(* Logix 5000 project; controller CIP vendor 1 type 14 code 106 rev 20.12; software revision 20.06; part 6 of 13 *)
(* tags used below, declared in another part *)
   Alarm_Ack : INT[8];
   Alarm_Ack_All_PB : BOOL;
   Alarm_Present : INT[8];
   Alarm_Remote_Ack_All : BOOL;
   Alarm_Status_Reset : BOOL;
   Bit : BOOL[128];
   IN_N7_100_199 : INT[100];
   Level_Bits : BOOL[32];
   Level_Timers : TIMER[20];
   Message_Index : ALIAS FOR Integer[30];
   Message_Present : INT[4];
   Message_SEQ : DINT[101];
   MOA_Status : DINT[10];
   One_Shot : BOOL[128];
   OpCode_Pin : DINT[5];
   Panelview : INT[40];
   PID1 : PID;
   PID2 : PID;
   PID3 : PID;
   PID3_Timer : TIMER[4];
   PID_Timer : TIMER[5];
   PV_Message : DINT[3];
   Recipe : RECIPE[41];
   Timer : TIMER[99];
   Timer_Chem1_Pump : TIMER[7];
   Timer_Chem2_Pump : TIMER[7];
   WashChamberDoorGasketCTRL : DINT;
(* MainProgram, continued *)

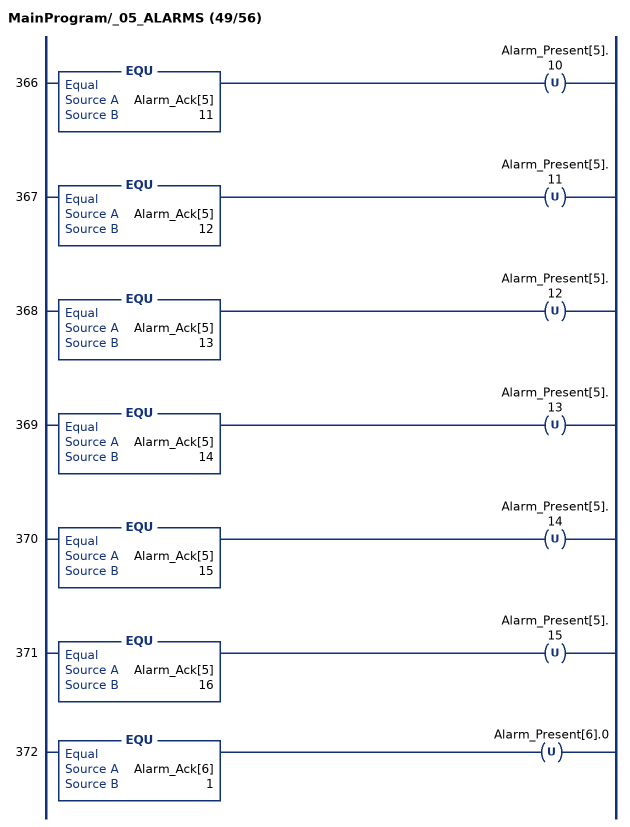
   [picture p91: MainProgram/_05_ALARMS rungs 366-372]
   366: EQU(Alarm_Ack[5],11)OTU(Alarm_Present[5].10);
   367: EQU(Alarm_Ack[5],12)OTU(Alarm_Present[5].11);
   368: EQU(Alarm_Ack[5],13)OTU(Alarm_Present[5].12);
   369: EQU(Alarm_Ack[5],14)OTU(Alarm_Present[5].13);
   370: EQU(Alarm_Ack[5],15)OTU(Alarm_Present[5].14);
   371: EQU(Alarm_Ack[5],16)OTU(Alarm_Present[5].15);
   372: EQU(Alarm_Ack[6],1)OTU(Alarm_Present[6].0);
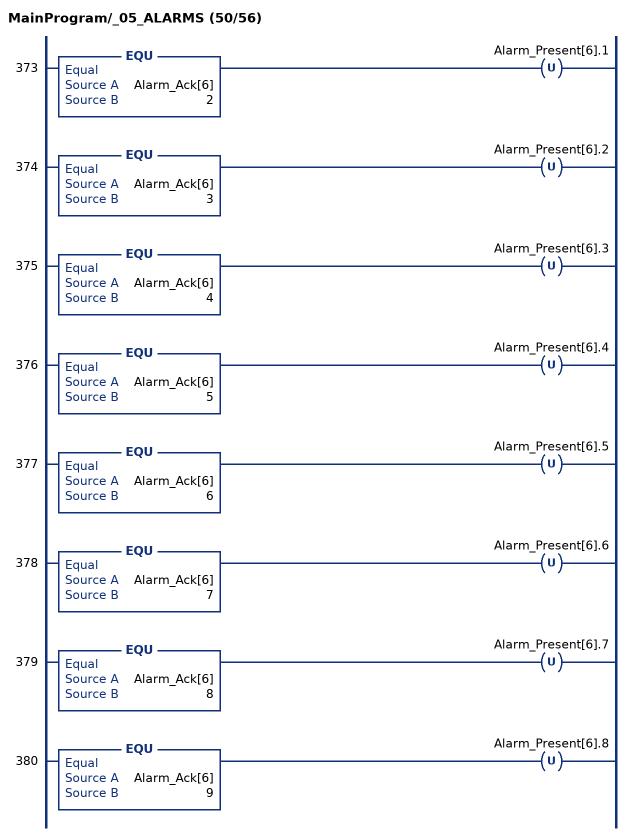
   373: EQU(Alarm_Ack[6],2)OTU(Alarm_Present[6].1);
   374: EQU(Alarm_Ack[6],3)OTU(Alarm_Present[6].2);
   375: EQU(Alarm_Ack[6],4)OTU(Alarm_Present[6].3);
   376: EQU(Alarm_Ack[6],5)OTU(Alarm_Present[6].4);
   377: EQU(Alarm_Ack[6],6)OTU(Alarm_Present[6].5);
   378: EQU(Alarm_Ack[6],7)OTU(Alarm_Present[6].6);
   379: EQU(Alarm_Ack[6],8)OTU(Alarm_Present[6].7);
   380: EQU(Alarm_Ack[6],9)OTU(Alarm_Present[6].8);
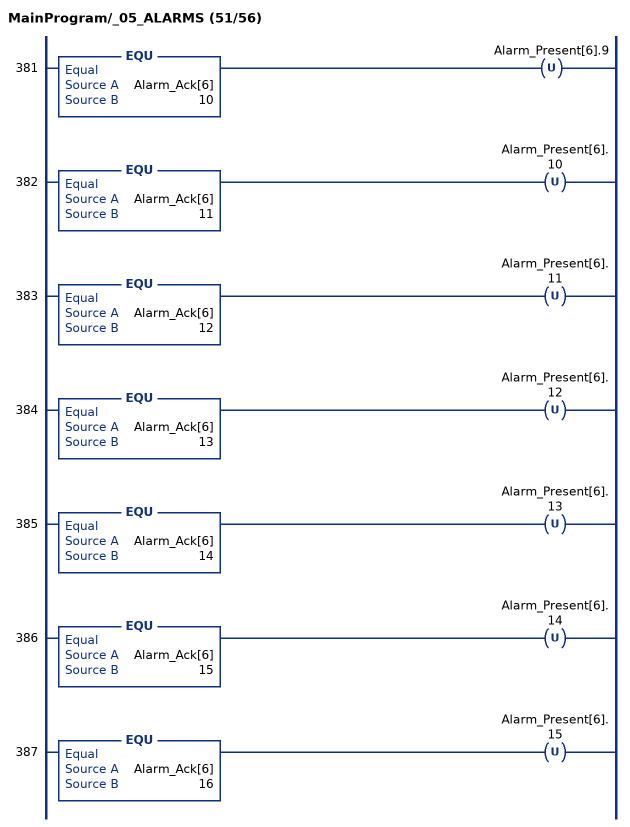
   381: EQU(Alarm_Ack[6],10)OTU(Alarm_Present[6].9);
   382: EQU(Alarm_Ack[6],11)OTU(Alarm_Present[6].10);
   383: EQU(Alarm_Ack[6],12)OTU(Alarm_Present[6].11);
   384: EQU(Alarm_Ack[6],13)OTU(Alarm_Present[6].12);
   385: EQU(Alarm_Ack[6],14)OTU(Alarm_Present[6].13);
   386: EQU(Alarm_Ack[6],15)OTU(Alarm_Present[6].14);
   387: EQU(Alarm_Ack[6],16)OTU(Alarm_Present[6].15);
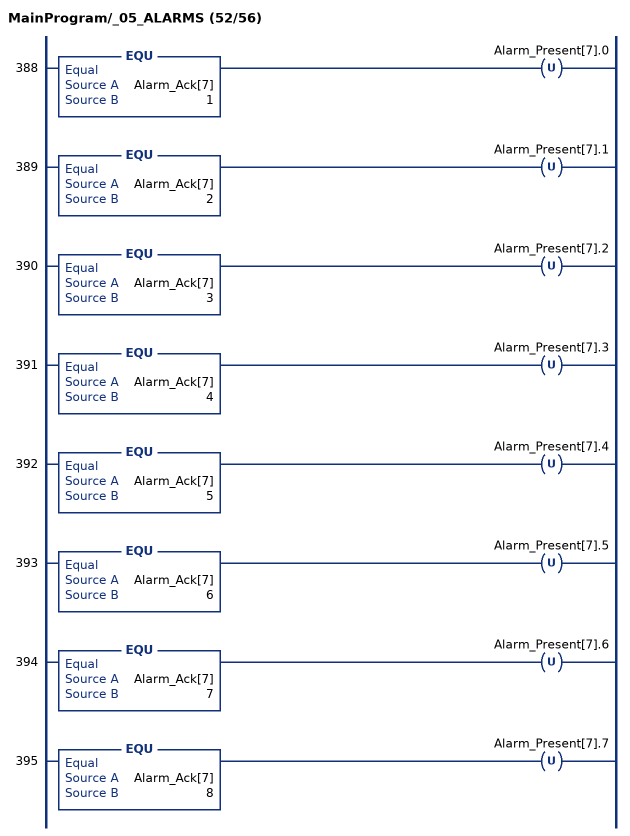
   388: EQU(Alarm_Ack[7],1)OTU(Alarm_Present[7].0);
   389: EQU(Alarm_Ack[7],2)OTU(Alarm_Present[7].1);
   390: EQU(Alarm_Ack[7],3)OTU(Alarm_Present[7].2);
   391: EQU(Alarm_Ack[7],4)OTU(Alarm_Present[7].3);
   392: EQU(Alarm_Ack[7],5)OTU(Alarm_Present[7].4);
   393: EQU(Alarm_Ack[7],6)OTU(Alarm_Present[7].5);
   394: EQU(Alarm_Ack[7],7)OTU(Alarm_Present[7].6);
   395: EQU(Alarm_Ack[7],8)OTU(Alarm_Present[7].7);
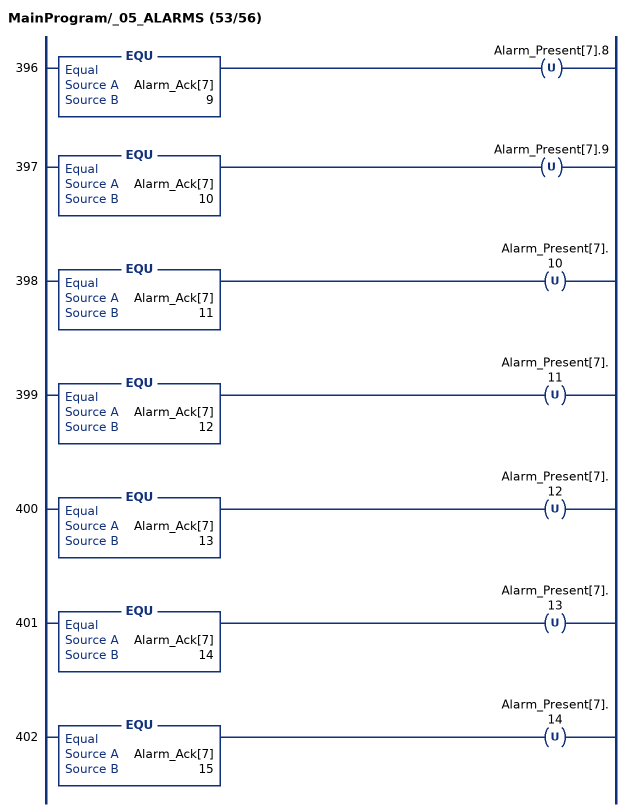
   396: EQU(Alarm_Ack[7],9)OTU(Alarm_Present[7].8);
   397: EQU(Alarm_Ack[7],10)OTU(Alarm_Present[7].9);
   398: EQU(Alarm_Ack[7],11)OTU(Alarm_Present[7].10);
   399: EQU(Alarm_Ack[7],12)OTU(Alarm_Present[7].11);
   400: EQU(Alarm_Ack[7],13)OTU(Alarm_Present[7].12);
   401: EQU(Alarm_Ack[7],14)OTU(Alarm_Present[7].13);
   402: EQU(Alarm_Ack[7],15)OTU(Alarm_Present[7].14);
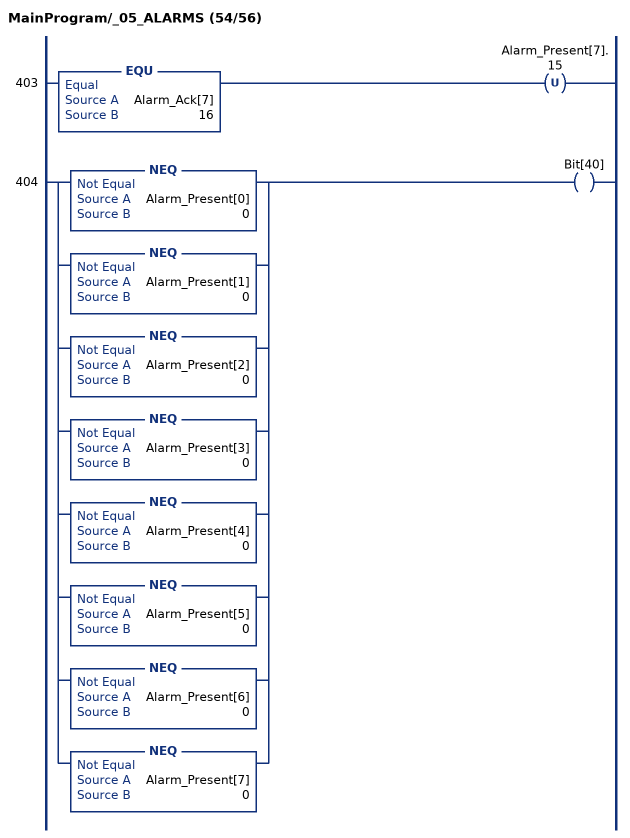
   403: EQU(Alarm_Ack[7],16)OTU(Alarm_Present[7].15);
   404: [NEQ(Alarm_Present[0],0) ,NEQ(Alarm_Present[1],0) ,NEQ(Alarm_Present[2],0) ,NEQ(Alarm_Present[3],0) ,NEQ(Alarm_Present[4],0) ,NEQ(Alarm_Present[5],0) ,NEQ(Alarm_Present[6],0) ,NEQ(Alarm_Present[7],0) ]OTE(Bit[40]);
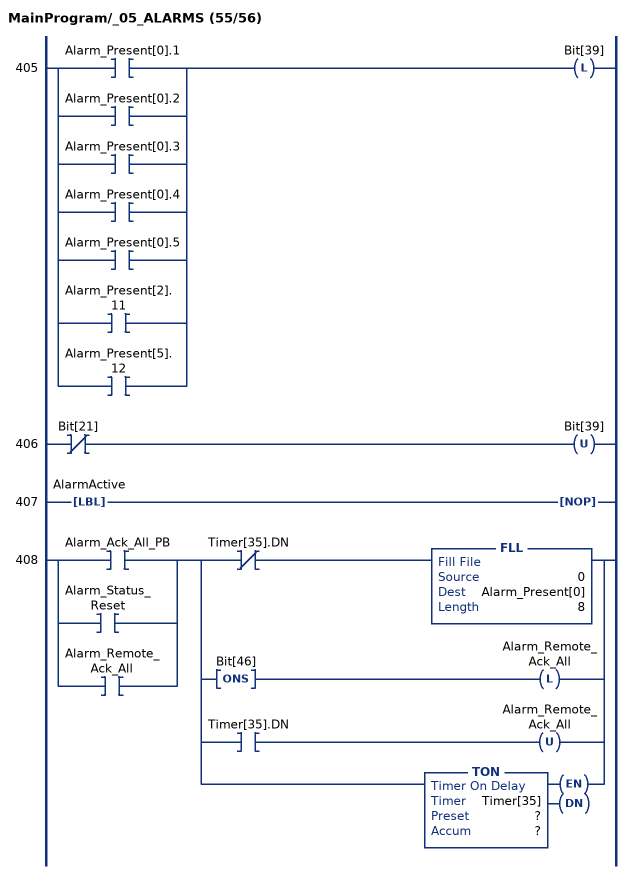
   405: [XIC(Alarm_Present[0].1) ,XIC(Alarm_Present[0].2) ,XIC(Alarm_Present[0].3) ,XIC(Alarm_Present[0].4) ,XIC(Alarm_Present[0].5) ,XIC(Alarm_Present[2].11) ,XIC(Alarm_Present[5].12) ]OTL(Bit[39]);
   406: XIO(Bit[21])OTU(Bit[39]);
   407: LBL(AlarmActive)NOP();
   408: [XIC(Alarm_Ack_All_PB) ,XIC(Alarm_Status_Reset) ,XIC(Alarm_Remote_Ack_All) ][XIO(Timer[35].DN) FLL(0,Alarm_Present[0],8) ,ONS(Bit[46]) OTL(Alarm_Remote_Ack_All) ,XIC(Timer[35].DN) OTU(Alarm_Remote_Ack_All) ,TON(Timer[35],?,?) ];
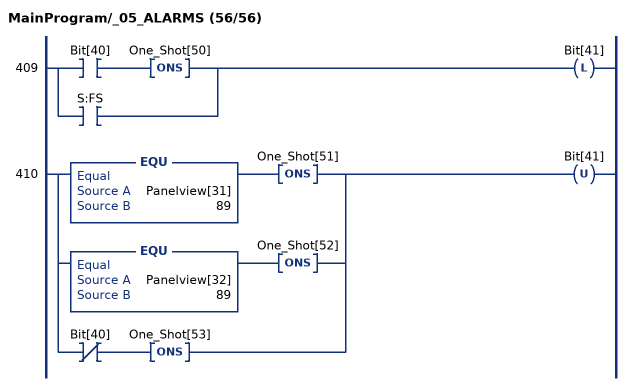
   409: [XIC(Bit[40]) ONS(One_Shot[50]) ,XIC(S:FS) ]OTL(Bit[41]);
   410: [EQU(Panelview[31],89) ONS(One_Shot[51]) ,EQU(Panelview[32],89) ONS(One_Shot[52]) ,XIO(Bit[40]) ONS(One_Shot[53]) ]OTU(Bit[41]);
END_ROUTINE

ROUTINE _05_MESSAGES   (* ladder *)
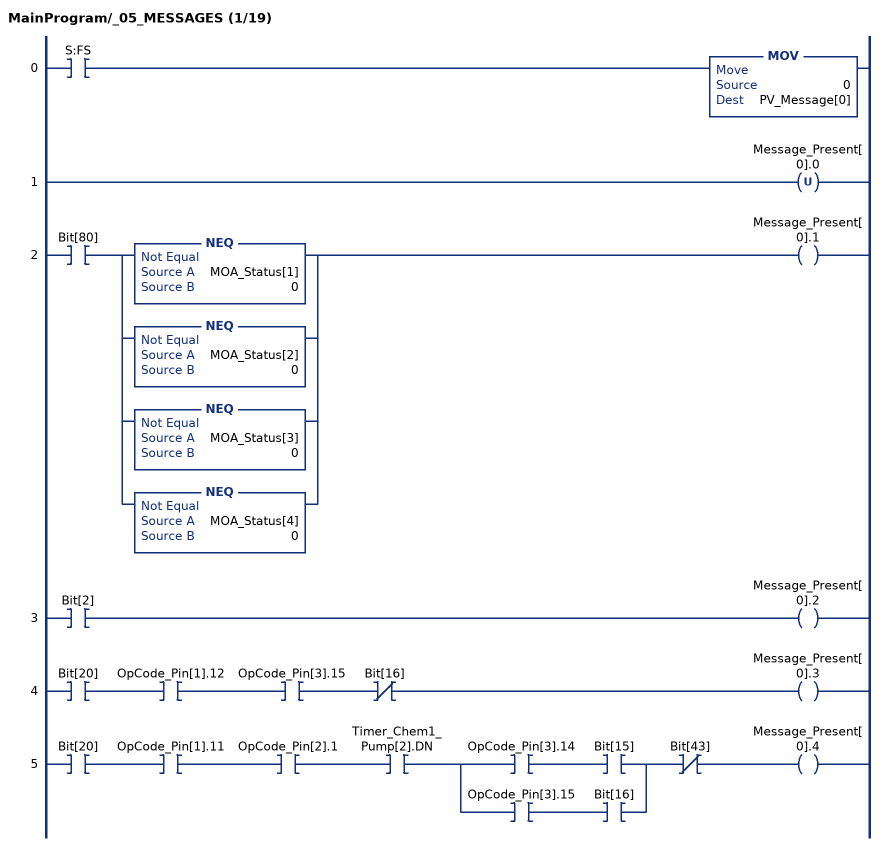
   0: XIC(S:FS)MOV(0,PV_Message[0]);
   1: OTU(Message_Present[0].0);
   2: XIC(Bit[80])[NEQ(MOA_Status[1],0) ,NEQ(MOA_Status[2],0) ,NEQ(MOA_Status[3],0) ,NEQ(MOA_Status[4],0) ]OTE(Message_Present[0].1);
   3: XIC(Bit[2])OTE(Message_Present[0].2);
   4: XIC(Bit[20])XIC(OpCode_Pin[1].12)XIC(OpCode_Pin[3].15)XIO(Bit[16])OTE(Message_Present[0].3);
   5: XIC(Bit[20])XIC(OpCode_Pin[1].11)XIC(OpCode_Pin[2].1)XIC(Timer_Chem1_Pump[2].DN)[XIC(OpCode_Pin[3].14) XIC(Bit[15]) ,XIC(OpCode_Pin[3].15) XIC(Bit[16]) ]XIO(Bit[43])OTE(Message_Present[0].4);
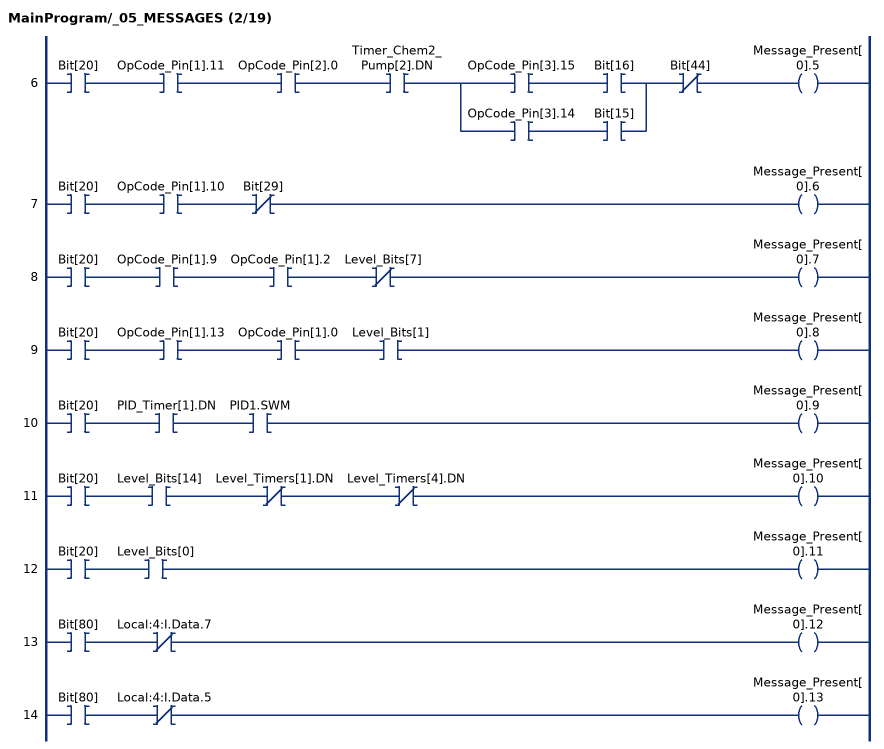
   6: XIC(Bit[20])XIC(OpCode_Pin[1].11)XIC(OpCode_Pin[2].0)XIC(Timer_Chem2_Pump[2].DN)[XIC(OpCode_Pin[3].15) XIC(Bit[16]) ,XIC(OpCode_Pin[3].14) XIC(Bit[15]) ]XIO(Bit[44])OTE(Message_Present[0].5);
   7: XIC(Bit[20])XIC(OpCode_Pin[1].10)XIO(Bit[29])OTE(Message_Present[0].6);
   8: XIC(Bit[20])XIC(OpCode_Pin[1].9)XIC(OpCode_Pin[1].2)XIO(Level_Bits[7])OTE(Message_Present[0].7);
   9: XIC(Bit[20])XIC(OpCode_Pin[1].13)XIC(OpCode_Pin[1].0)XIC(Level_Bits[1])OTE(Message_Present[0].8);
   10: XIC(Bit[20])XIC(PID_Timer[1].DN)XIC(PID1.SWM)OTE(Message_Present[0].9);
   11: XIC(Bit[20])XIC(Level_Bits[14])XIO(Level_Timers[1].DN)XIO(Level_Timers[4].DN)OTE(Message_Present[0].10);
   12: XIC(Bit[20])XIC(Level_Bits[0])OTE(Message_Present[0].11);
   13: XIC(Bit[80])XIO(Local:4:I.Data.7)OTE(Message_Present[0].12);
   14: XIC(Bit[80])XIO(Local:4:I.Data.5)OTE(Message_Present[0].13);
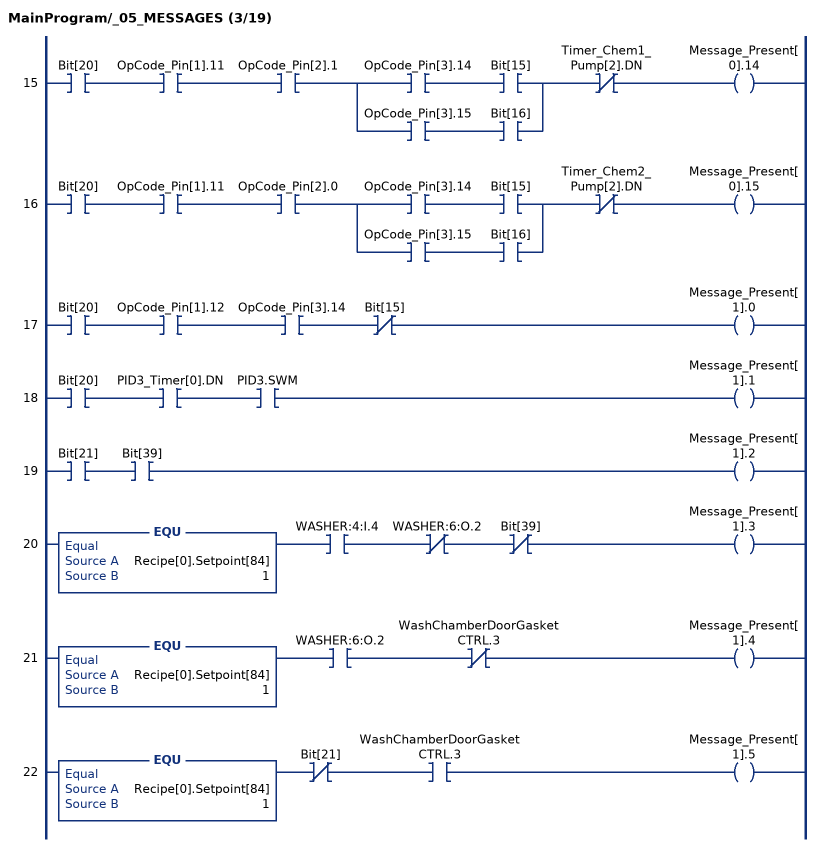
   15: XIC(Bit[20])XIC(OpCode_Pin[1].11)XIC(OpCode_Pin[2].1)[XIC(OpCode_Pin[3].14) XIC(Bit[15]) ,XIC(OpCode_Pin[3].15) XIC(Bit[16]) ]XIO(Timer_Chem1_Pump[2].DN)OTE(Message_Present[0].14);
   16: XIC(Bit[20])XIC(OpCode_Pin[1].11)XIC(OpCode_Pin[2].0)[XIC(OpCode_Pin[3].14) XIC(Bit[15]) ,XIC(OpCode_Pin[3].15) XIC(Bit[16]) ]XIO(Timer_Chem2_Pump[2].DN)OTE(Message_Present[0].15);
   17: XIC(Bit[20])XIC(OpCode_Pin[1].12)XIC(OpCode_Pin[3].14)XIO(Bit[15])OTE(Message_Present[1].0);
   18: XIC(Bit[20])XIC(PID3_Timer[0].DN)XIC(PID3.SWM)OTE(Message_Present[1].1);
   19: XIC(Bit[21])XIC(Bit[39])OTE(Message_Present[1].2);
   20: EQU(Recipe[0].Setpoint[84],1)XIC(WASHER:4:I.4)XIO(WASHER:6:O.2)XIO(Bit[39])OTE(Message_Present[1].3);
   21: EQU(Recipe[0].Setpoint[84],1)XIC(WASHER:6:O.2)XIO(WashChamberDoorGasketCTRL.3)OTE(Message_Present[1].4);
   22: EQU(Recipe[0].Setpoint[84],1)XIO(Bit[21])XIC(WashChamberDoorGasketCTRL.3)OTE(Message_Present[1].5);
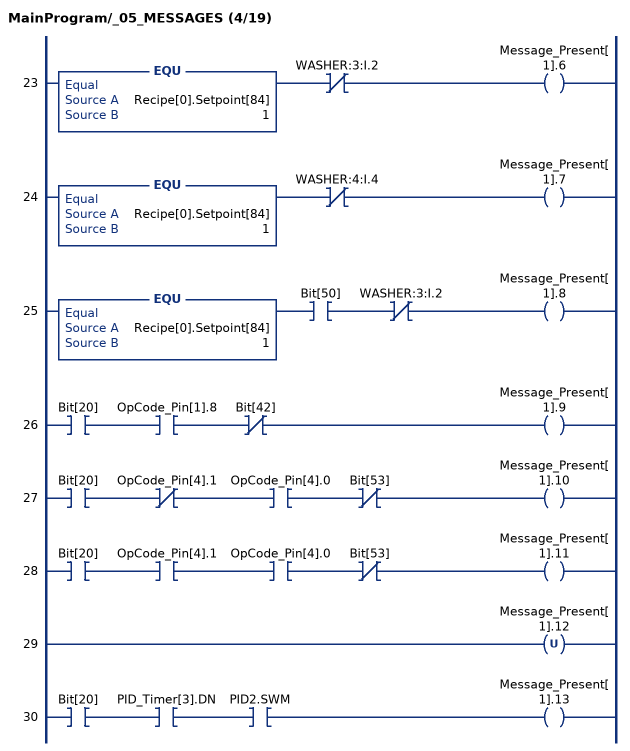
   23: EQU(Recipe[0].Setpoint[84],1)XIO(WASHER:3:I.2)OTE(Message_Present[1].6);
   24: EQU(Recipe[0].Setpoint[84],1)XIO(WASHER:4:I.4)OTE(Message_Present[1].7);
   25: EQU(Recipe[0].Setpoint[84],1)XIC(Bit[50])XIO(WASHER:3:I.2)OTE(Message_Present[1].8);
   26: XIC(Bit[20])XIC(OpCode_Pin[1].8)XIO(Bit[42])OTE(Message_Present[1].9);
   27: XIC(Bit[20])XIO(OpCode_Pin[4].1)XIC(OpCode_Pin[4].0)XIO(Bit[53])OTE(Message_Present[1].10);
   28: XIC(Bit[20])XIC(OpCode_Pin[4].1)XIC(OpCode_Pin[4].0)XIO(Bit[53])OTE(Message_Present[1].11);
   29: OTU(Message_Present[1].12);
   30: XIC(Bit[20])XIC(PID_Timer[3].DN)XIC(PID2.SWM)OTE(Message_Present[1].13);
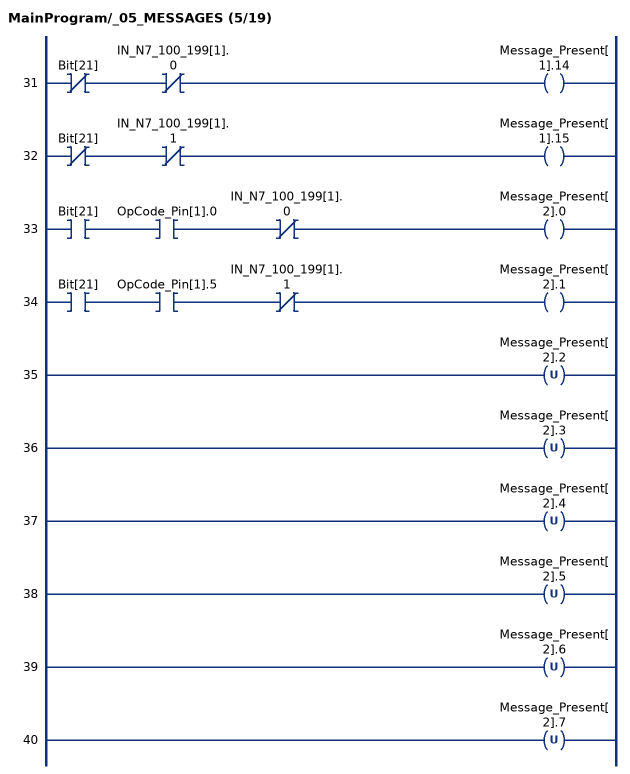
   31: XIO(Bit[21])XIO(IN_N7_100_199[1].0)OTE(Message_Present[1].14);
   32: XIO(Bit[21])XIO(IN_N7_100_199[1].1)OTE(Message_Present[1].15);
   33: XIC(Bit[21])XIC(OpCode_Pin[1].0)XIO(IN_N7_100_199[1].0)OTE(Message_Present[2].0);
   34: XIC(Bit[21])XIC(OpCode_Pin[1].5)XIO(IN_N7_100_199[1].1)OTE(Message_Present[2].1);
   35: OTU(Message_Present[2].2);
   36: OTU(Message_Present[2].3);
   37: OTU(Message_Present[2].4);
   38: OTU(Message_Present[2].5);
   39: OTU(Message_Present[2].6);
   40: OTU(Message_Present[2].7);
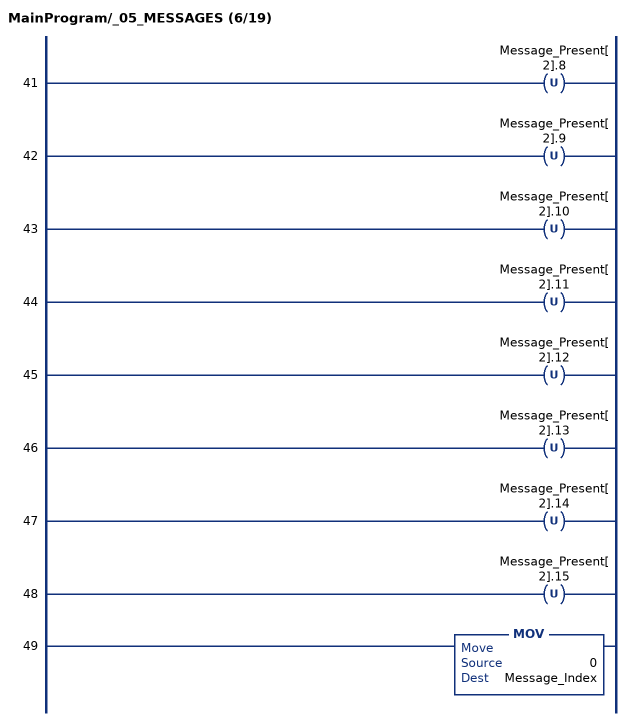
   41: OTU(Message_Present[2].8);
   42: OTU(Message_Present[2].9);
   43: OTU(Message_Present[2].10);
   44: OTU(Message_Present[2].11);
   45: OTU(Message_Present[2].12);
   46: OTU(Message_Present[2].13);
   47: OTU(Message_Present[2].14);
   48: OTU(Message_Present[2].15);
   49: MOV(0,Message_Index);
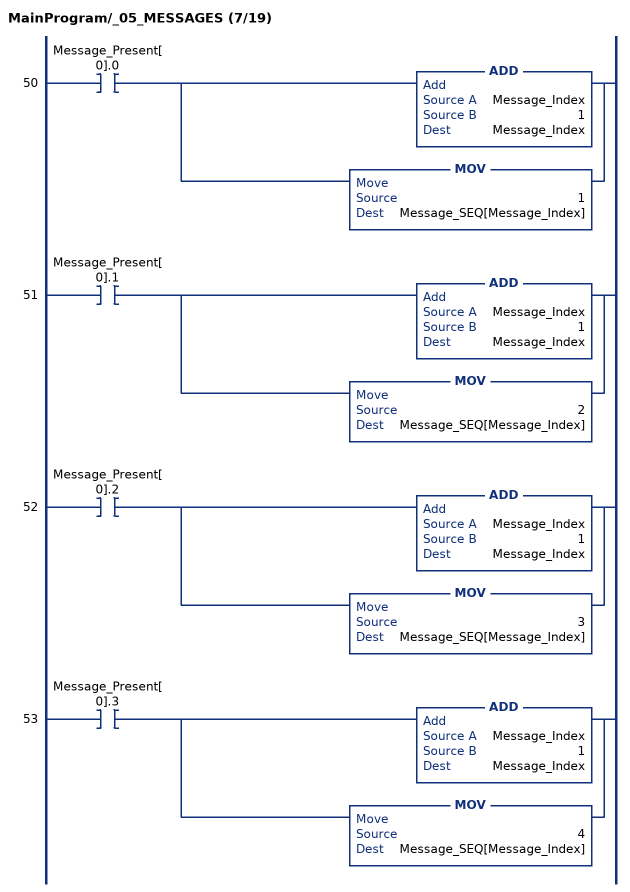
   50: XIC(Message_Present[0].0)[ADD(Message_Index,1,Message_Index) ,MOV(1,Message_SEQ[Message_Index]) ];
   51: XIC(Message_Present[0].1)[ADD(Message_Index,1,Message_Index) ,MOV(2,Message_SEQ[Message_Index]) ];
   52: XIC(Message_Present[0].2)[ADD(Message_Index,1,Message_Index) ,MOV(3,Message_SEQ[Message_Index]) ];
   53: XIC(Message_Present[0].3)[ADD(Message_Index,1,Message_Index) ,MOV(4,Message_SEQ[Message_Index]) ];
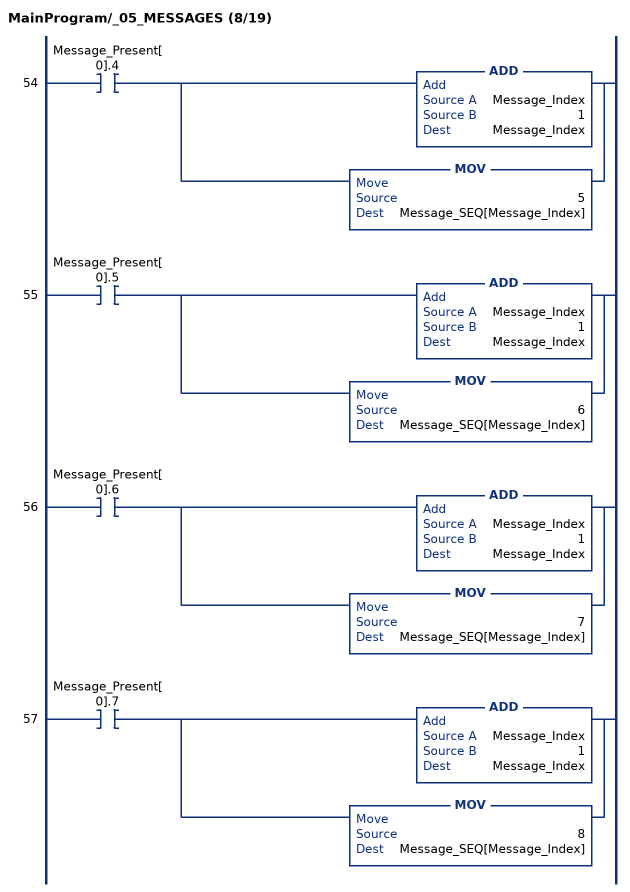
   54: XIC(Message_Present[0].4)[ADD(Message_Index,1,Message_Index) ,MOV(5,Message_SEQ[Message_Index]) ];
   55: XIC(Message_Present[0].5)[ADD(Message_Index,1,Message_Index) ,MOV(6,Message_SEQ[Message_Index]) ];
   56: XIC(Message_Present[0].6)[ADD(Message_Index,1,Message_Index) ,MOV(7,Message_SEQ[Message_Index]) ];
   57: XIC(Message_Present[0].7)[ADD(Message_Index,1,Message_Index) ,MOV(8,Message_SEQ[Message_Index]) ];
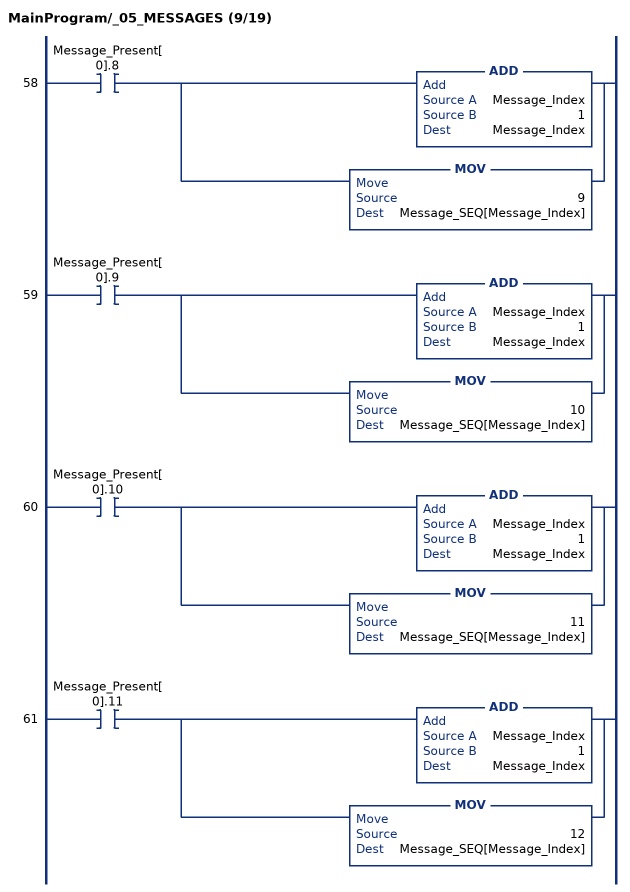
   58: XIC(Message_Present[0].8)[ADD(Message_Index,1,Message_Index) ,MOV(9,Message_SEQ[Message_Index]) ];
   59: XIC(Message_Present[0].9)[ADD(Message_Index,1,Message_Index) ,MOV(10,Message_SEQ[Message_Index]) ];
   60: XIC(Message_Present[0].10)[ADD(Message_Index,1,Message_Index) ,MOV(11,Message_SEQ[Message_Index]) ];
   61: XIC(Message_Present[0].11)[ADD(Message_Index,1,Message_Index) ,MOV(12,Message_SEQ[Message_Index]) ];
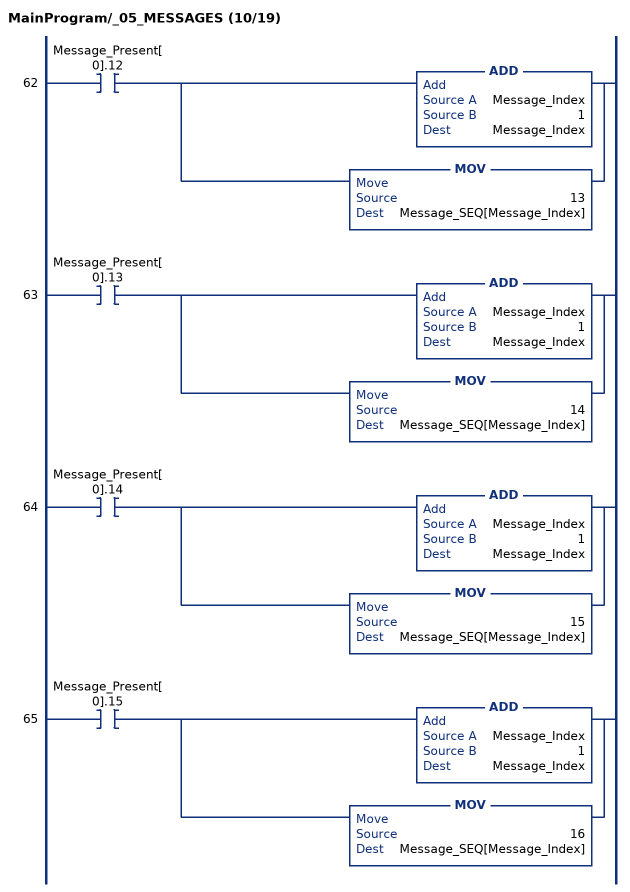
   62: XIC(Message_Present[0].12)[ADD(Message_Index,1,Message_Index) ,MOV(13,Message_SEQ[Message_Index]) ];
   63: XIC(Message_Present[0].13)[ADD(Message_Index,1,Message_Index) ,MOV(14,Message_SEQ[Message_Index]) ];
   64: XIC(Message_Present[0].14)[ADD(Message_Index,1,Message_Index) ,MOV(15,Message_SEQ[Message_Index]) ];
   65: XIC(Message_Present[0].15)[ADD(Message_Index,1,Message_Index) ,MOV(16,Message_SEQ[Message_Index]) ];
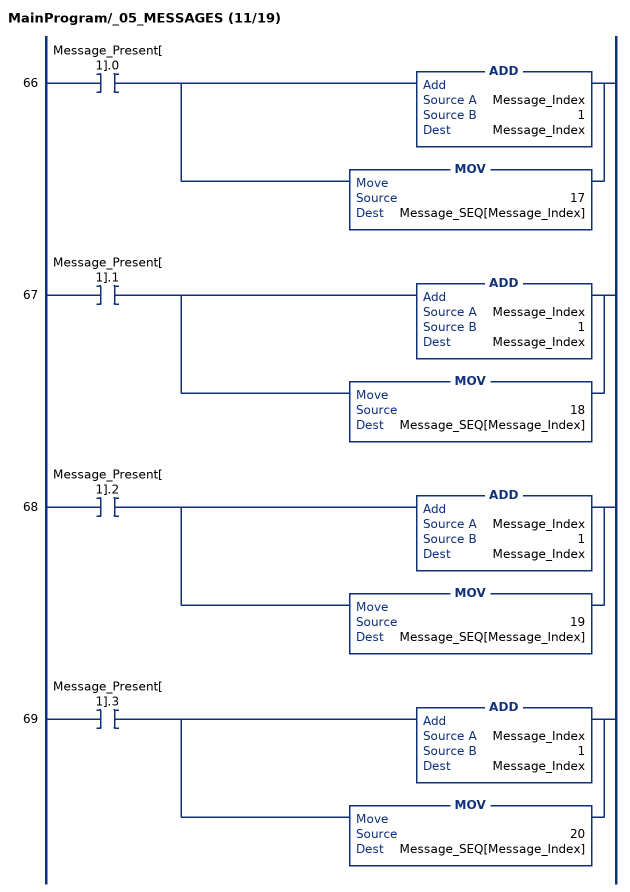
   66: XIC(Message_Present[1].0)[ADD(Message_Index,1,Message_Index) ,MOV(17,Message_SEQ[Message_Index]) ];
   67: XIC(Message_Present[1].1)[ADD(Message_Index,1,Message_Index) ,MOV(18,Message_SEQ[Message_Index]) ];
   68: XIC(Message_Present[1].2)[ADD(Message_Index,1,Message_Index) ,MOV(19,Message_SEQ[Message_Index]) ];
   69: XIC(Message_Present[1].3)[ADD(Message_Index,1,Message_Index) ,MOV(20,Message_SEQ[Message_Index]) ];
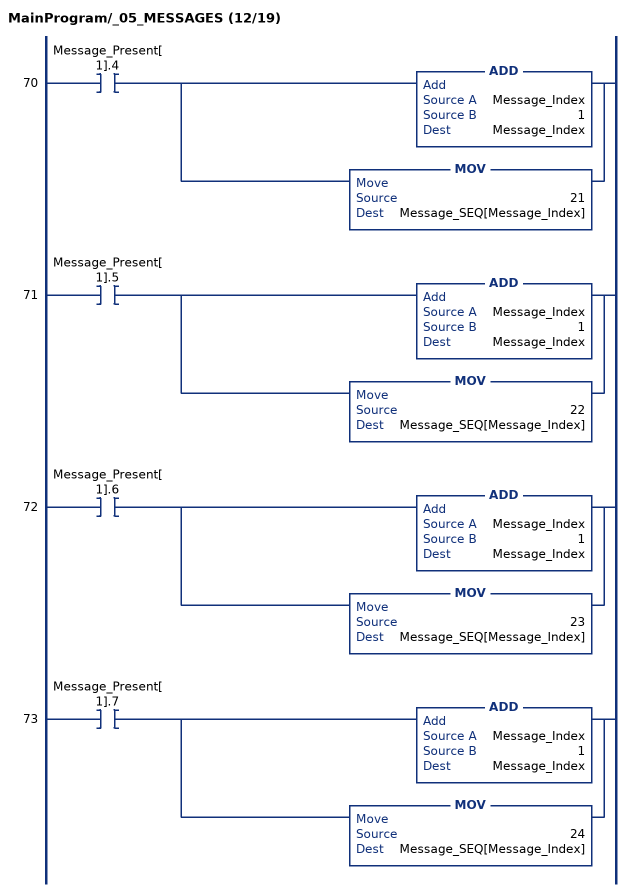
   70: XIC(Message_Present[1].4)[ADD(Message_Index,1,Message_Index) ,MOV(21,Message_SEQ[Message_Index]) ];
   71: XIC(Message_Present[1].5)[ADD(Message_Index,1,Message_Index) ,MOV(22,Message_SEQ[Message_Index]) ];
   72: XIC(Message_Present[1].6)[ADD(Message_Index,1,Message_Index) ,MOV(23,Message_SEQ[Message_Index]) ];
   73: XIC(Message_Present[1].7)[ADD(Message_Index,1,Message_Index) ,MOV(24,Message_SEQ[Message_Index]) ];
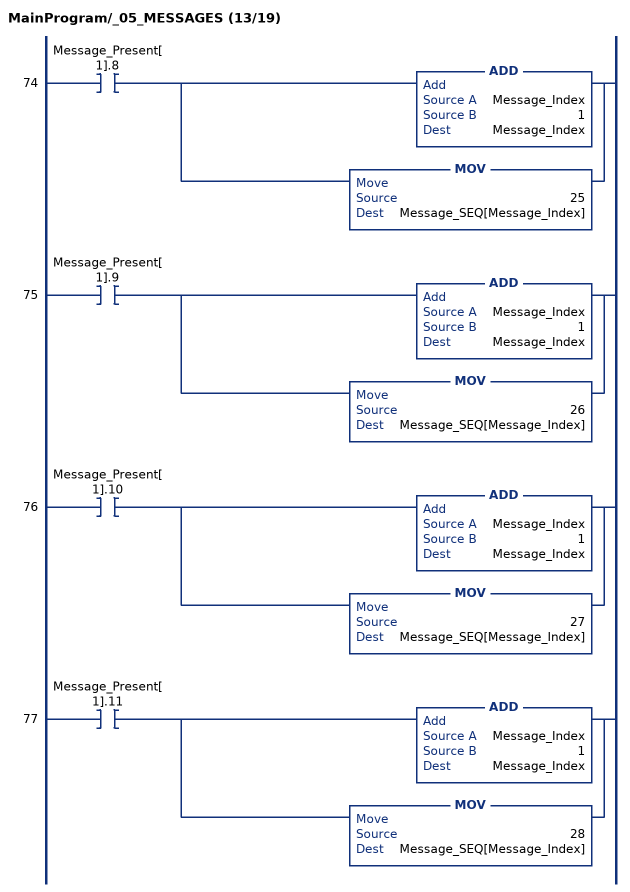
   74: XIC(Message_Present[1].8)[ADD(Message_Index,1,Message_Index) ,MOV(25,Message_SEQ[Message_Index]) ];
   75: XIC(Message_Present[1].9)[ADD(Message_Index,1,Message_Index) ,MOV(26,Message_SEQ[Message_Index]) ];
   76: XIC(Message_Present[1].10)[ADD(Message_Index,1,Message_Index) ,MOV(27,Message_SEQ[Message_Index]) ];
   77: XIC(Message_Present[1].11)[ADD(Message_Index,1,Message_Index) ,MOV(28,Message_SEQ[Message_Index]) ];
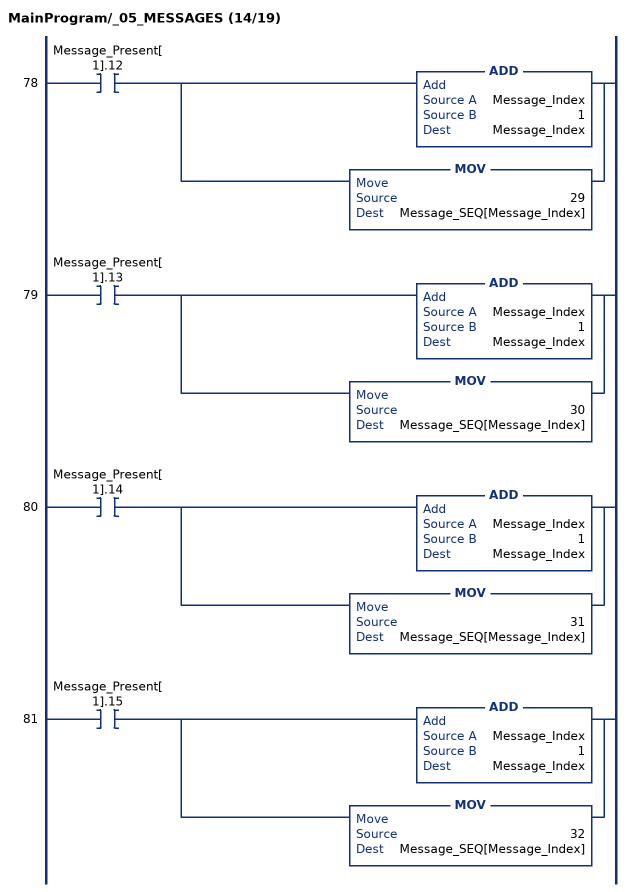
   78: XIC(Message_Present[1].12)[ADD(Message_Index,1,Message_Index) ,MOV(29,Message_SEQ[Message_Index]) ];
   79: XIC(Message_Present[1].13)[ADD(Message_Index,1,Message_Index) ,MOV(30,Message_SEQ[Message_Index]) ];
   80: XIC(Message_Present[1].14)[ADD(Message_Index,1,Message_Index) ,MOV(31,Message_SEQ[Message_Index]) ];
   81: XIC(Message_Present[1].15)[ADD(Message_Index,1,Message_Index) ,MOV(32,Message_SEQ[Message_Index]) ];
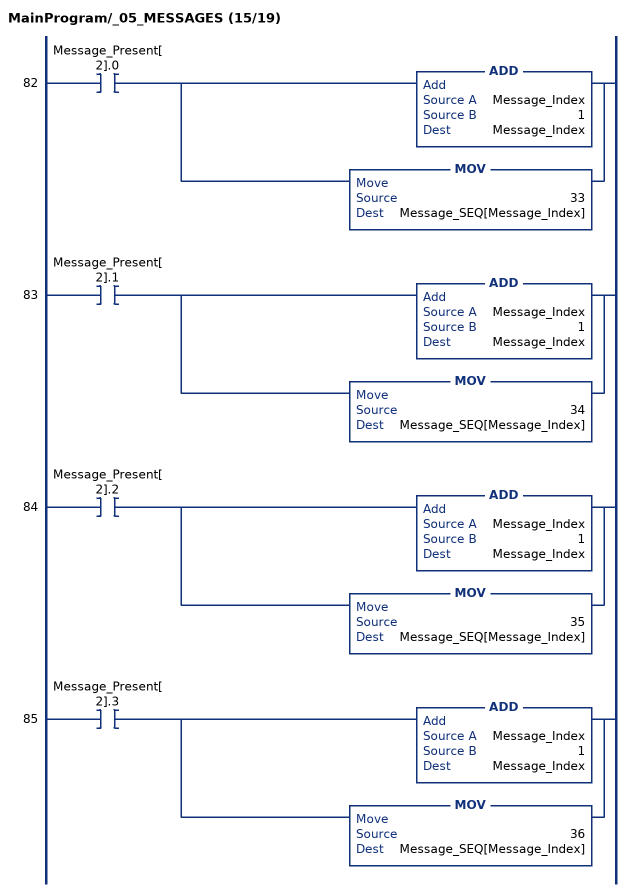
   82: XIC(Message_Present[2].0)[ADD(Message_Index,1,Message_Index) ,MOV(33,Message_SEQ[Message_Index]) ];
   83: XIC(Message_Present[2].1)[ADD(Message_Index,1,Message_Index) ,MOV(34,Message_SEQ[Message_Index]) ];
   84: XIC(Message_Present[2].2)[ADD(Message_Index,1,Message_Index) ,MOV(35,Message_SEQ[Message_Index]) ];
   85: XIC(Message_Present[2].3)[ADD(Message_Index,1,Message_Index) ,MOV(36,Message_SEQ[Message_Index]) ];
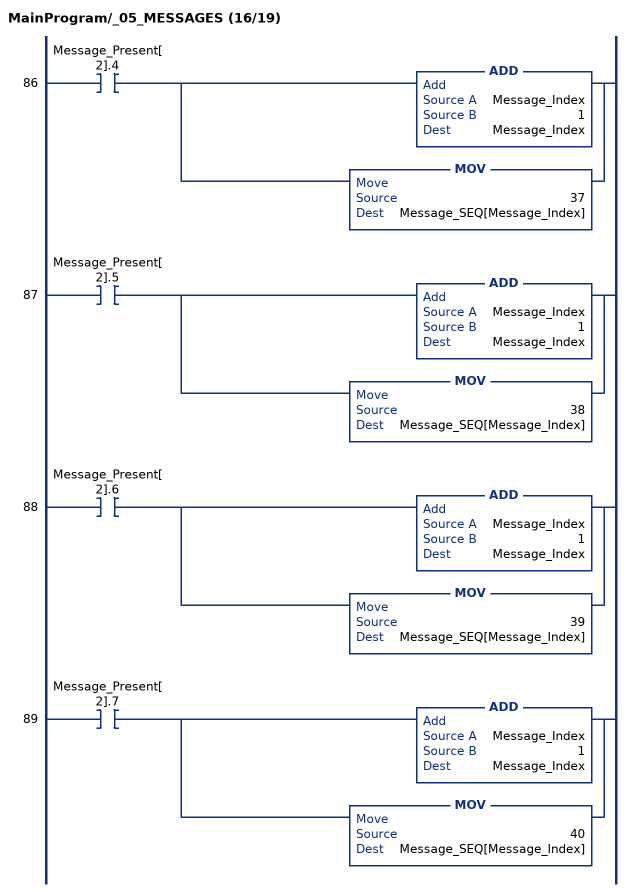
   86: XIC(Message_Present[2].4)[ADD(Message_Index,1,Message_Index) ,MOV(37,Message_SEQ[Message_Index]) ];
   87: XIC(Message_Present[2].5)[ADD(Message_Index,1,Message_Index) ,MOV(38,Message_SEQ[Message_Index]) ];
   88: XIC(Message_Present[2].6)[ADD(Message_Index,1,Message_Index) ,MOV(39,Message_SEQ[Message_Index]) ];
   89: XIC(Message_Present[2].7)[ADD(Message_Index,1,Message_Index) ,MOV(40,Message_SEQ[Message_Index]) ];
